(* Basic Input Output Example *)

PROGRAM main
  VAR
    Input AT %IX0.0 : BOOL;
    Output AT %QX0.0 : BOOL; (* Output Coil 1 *)
  END_VAR

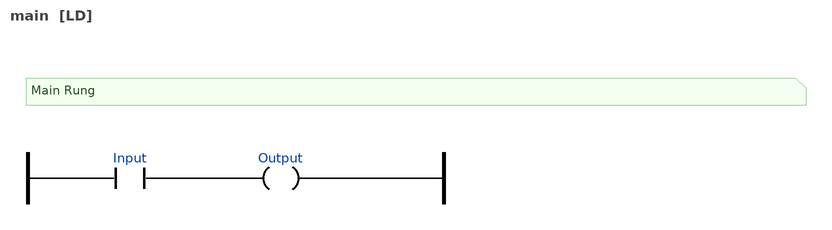
(* LD diagram, written out as Structured Text *)
(* Main Rung *)
Output := Input;
END_PROGRAM
